Universal Robots URScript: ConfProg.script

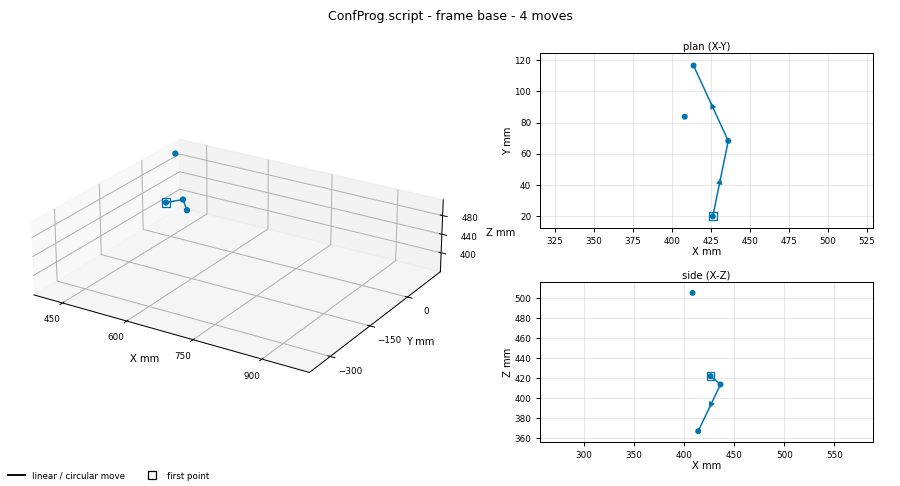
[picture p0: tool path of ConfProg.script in frame base, 4 of 6 moves have a stored position in this frame; points joined in program order, loops and branches not executed]
def ConfProg():
  # Global parameters:
  global speed_ms    = 0.250
  global speed_rads  = 0.750
  global accel_mss   = 1.200
  global accel_radss = 1.200
  global blend_radius_m = 0.000

  #--------------------------
  # Add any default subprograms here
  # For example, to drive a gripper as a program call:
  # def Gripper_Open():
  #   ...
  # end
  #
  # Example to drive a spray gun:
  def SprayOn(value):
    # use the value as an output:
    DO_SPRAY = 5
    if value == 0:
      set_standard_digital_out(DO_SPRAY, False)
    else:
      set_standard_digital_out(DO_SPRAY, True)
    end
  end

  # Example to synchronize 2
  def Synchronize():
    # Use the following digital output to signal the state of the robot:
    DO_SYNC = 1

    # Use the following digital input to get the state of another robot:
    DI_SYNC = 1

    if (get_standard_digital_out(DO_SYNC) == get_standard_digital_in(DI_SYNC)):
      set_standard_digital_out(DO_SYNC, not (get_standard_digital_out(DI_SYNC)))
      sleep(0.1)
      thread Thread_wait_1():
        while (True):
          sleep(0.01)
        end
      end
      if (get_standard_digital_out(DO_SYNC) != get_standard_digital_in(DI_SYNC)):
        global thread_handler_1=run Thread_wait_1()
        while (get_standard_digital_out(DO_SYNC) != get_standard_digital_in(DI_SYNC)):
          sync()
        end
        kill thread_handler_1
      end
    else:
      if (get_standard_digital_out(DO_SYNC) != get_standard_digital_in(DI_SYNC)):
        set_standard_digital_out(DO_SYNC, not (get_standard_digital_out(DO_SYNC)))
      end
    end
  end

  #
  # Example to move an external axis
  def MoveAxis(value):
    # use the value as an output:
    DO_AXIS_1 = 1
    DI_AXIS_1 = 1
    if value <= 0:
      set_standard_digital_out(DO_AXIS_1, False)

      # Wait for digital input to change state
      #while (get_standard_digital_in(DI_AXIS_1) != False):
      #  sync()
      #end
    else:
      set_standard_digital_out(DO_AXIS_1, True)

      # Wait for digital input to change state
      #while (get_standard_digital_in(DI_AXIS_1) != True):
      #  sync()
      #end
    end
  end
  #--------------------------


  # Main program:
  # Program generated by RoboDK v6.0.7 for ABB IRB 120-3/0.6 on XX/XX/XXXX 18:00:00
  # Using nominal kinematics.
  # Using Ref. Frame S: p[1.234570, -0.098765, 0.050500, 0.000000, 0.000000, 0.523599]
  # set_reference(p[1.234570, -0.098765, 0.050500, 0.000000, 0.000000, 0.523599])
  # Using TCP Tool S: p[0.010000, 0.020000, 0.150000, 0.000000, 0.000000, 0.000000]
  set_tcp(p[0.010000, 0.020000, 0.150000, 0.000000, 0.000000, 0.000000])
  movel(p[0.426318, 0.020000, 0.422034, 0.138328, 2.253250, -0.296646],accel_mss,speed_ms,0,0.000)
  movel(p[0.436232, 0.068297, 0.413715, 0.138328, 2.253250, -0.296646],accel_mss,speed_ms,0,0.000)
  movel(p[0.414005, 0.116593, 0.367095, 0.138328, 2.253250, -0.296646],accel_mss,speed_ms,0,0.000)
  movej([0.174533, 0.349066, -0.523599, 0.698132, -0.872665, 1.047198],1.20000,0.75000,0,0.0000)
  movej([-2.967060, 0.785398, -0.785398, -2.967060, 1.570796, -3.124139],1.20000,0.75000,0,0.0000)
  # Circular move (R405.1 mm)
  movec(p[0.973908, -0.353337, 0.382202, -0.503745, 2.359457, 0.000119],p[0.408367, 0.083800, 0.505120, -0.487372, 1.445847, -0.747268],1.20000,0.25000,0.0000)
  # End of main program
end

ConfProg()
